Fanuc KAREL source: KO00145.KL

PROGRAM KO00145
%NOLOCKGROUP
VAR
  R: REAL
  CFG: CONFIG
  OUT: XYZWPR
  N: INTEGER
BEGIN
  N = 1
  R = 2.0
  CFG.CFG_FLIP = TRUE
  OUT = POS(R, R, R, R, N, R, CFG)
END KO00145
